Fanuc KAREL source: NC0062.KL

PROGRAM NC0062
%NOLOCKGROUP
ROUTINE R
VAR
  X : INTEGER
  I1 : INTEGER
BEGIN
  X = 1
  FOR I1 = 1 TO 2 DO
    X = X + 1
  ENDFOR
END R
BEGIN
  R
END NC0062
